// TIA Portal V17 program export: 0 tag tables, 0 data types, 0 data blocks, 2 code blocks (in call order from the OBs), 0 instance data blocks

ORGANIZATION_BLOCK "Main"   // OB1, LAD, ProgramCycle
TITLE = Programa principal
{ S7_Optimized_Access := 'TRUE' }
// Generado automáticamente con Claude Code + TIA Openness
   VAR_INPUT
      Initial_Call : Bool;   // Initial call of this OB
      Remanence : Bool;   // =True, if remanent data are available
   END_VAR
BEGIN

REGION Network 1: Motor 1
   // Llamada al bloque de arranque y paro con las entradas/salidas físicas
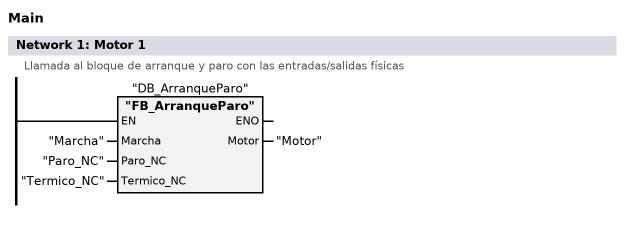
   RUNG wire#powerrail
      "DB_ArranqueParo"(Marcha := "Marcha", Paro_NC := "Paro_NC", Termico_NC := "Termico_NC", Motor => "Motor")
   END_RUNG
   // the same network as SCL:
   "DB_ArranqueParo"(Marcha := "Marcha", Paro_NC := "Paro_NC", Termico_NC := "Termico_NC", Motor => "Motor");   // "FB_ArranqueParo"
END_REGION
END_ORGANIZATION_BLOCK

FUNCTION_BLOCK "FB_ArranqueParo"   // FB1, LAD
TITLE = Arranque y paro de motor
{ S7_Optimized_Access := 'TRUE' }
// Generado automáticamente con Claude Code + TIA Openness
   VAR_INPUT
      Marcha : Bool;   // Pulsador de marcha (NA)
      Paro_NC : Bool;   // Pulsador de paro (NC)
      Termico_NC : Bool;   // Relé térmico (NC)
   END_VAR
   VAR_OUTPUT
      Motor : Bool;   // Orden al contactor del motor
   END_VAR
BEGIN

REGION Network 1: Arranque y paro con retención
   // Marcha arranca el motor y el propio contacto de Motor lo mantiene (retención). Paro o falla del térmico lo detienen. Paro dominante.
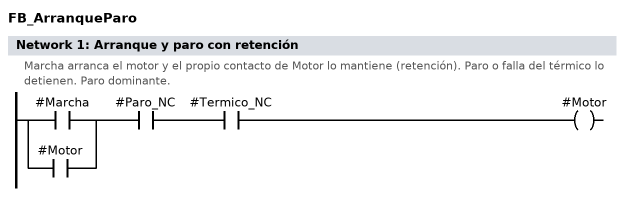
   RUNG wire#powerrail
      Contact( #Marcha )
      wire#w1
      Contact( #Paro_NC )
      Contact( #Termico_NC )
      Coil( #Motor )
   END_RUNG
   RUNG wire#powerrail
      Contact( #Motor )
   END_RUNG wire#w1
   // the same network as SCL:
   #Motor := (#Marcha OR #Motor) AND #Paro_NC AND #Termico_NC;
END_REGION
END_FUNCTION_BLOCK
